Yaskawa INFORM job: JOINTTA.JBI

/JOB
//NAME JOINTTA
//POS
///NPOS 11,0,0,0,0,0
///TOOL 1
///POSTYPE PULSE
///PULSE
C00000=10,20,-10,30,-45,60
C00001=18,24,-10,30,-45,60
C00002=18,24,-10,30,-45,60
C00003=10,20,-10,30,-45,60
C00004=18,24,-10,30,-45,60
C00005=10,20,-10,30,-45,60
C00006=18,24,-10,30,-45,60
C00007=18,24,-10,30,-45,60
C00008=10,20,-10,30,-45,60
C00009=18,24,-10,30,-45,60
C00010=10,20,-10,30,-45,60
//INST
///DATE 2026/10/26 01:18
///COMM Generated using RoboDK
///ATTR SC,RW
///GROUP1 RB1
NOP
'Program generated by Vertical
'Bot Studio for Motoman GP8 on
' 25/10/2026 12:00:00
'Using nominal kinematics.
'Using Frame 2 (targets wrt ba
'se):
'100.0,-50.0,20.0,0.0,0.0,30.0
'Tool 1 (Tool 1) should be clo
'se to:
'10.0,0.0,120.0,0.0,15.0,0.0
MOVJ C00000 VJ=50.00
MOVL C00001 V=100.0
MOVJ C00002 VJ=50.00
MOVL C00003 V=100.0
MOVL C00004 V=100.0
MOVJ C00005 VJ=50.00 PL=5
MOVL C00006 V=100.0 PL=5
MOVJ C00007 VJ=50.00 PL=5
MOVL C00008 V=100.0 PL=5
MOVL C00009 V=100.0 PL=5
MOVJ C00010 VJ=50.00
END
